Fanuc KAREL source: KT00522.KL

PROGRAM KT00522
%NOLOCKGROUP
VAR
  P1: XYZWPREXT
  P2: XYZWPR
  OUT: JOINTPOS
BEGIN
  P1.X = 1.0
    P2.Y = 2.0
  OUT = P1 : P2
END KT00522
